(* IEC 61131-3 sources: codesys-framework/txt/application/WeVe IO (library)/DigitalInput/FB_DigitalInput, 2 files *)

(* ---- Signals.prop.st ---- *)
PROPERTY Signals : SC_DigitalInputSignals

// --- BEGIN IMPLEMENTATION ---

// ----------- GET -----------
VAR
END_VAR

// -- BEGIN IMPLEMENTATION GET --
Signals := _scDISignals;

(* ---- SysPar.prop.st ---- *)
PROPERTY SysPar : SC_SystemParametersDigitalInput

// --- BEGIN IMPLEMENTATION ---

// ----------- SET -----------
VAR
END_VAR

// -- BEGIN IMPLEMENTATION SET --
_scSysPar := SysPar;
